(* IEC 61131-3 sources: codesys-framework/txt/application/WeVe IO (library)/Analog Input/FB_AnalogInput, 2 files *)

(* ---- Signals.prop.st ---- *)
PROPERTY Signals : SC_AnalogInputSignals

// --- BEGIN IMPLEMENTATION ---

// ----------- GET -----------
VAR
END_VAR

// -- BEGIN IMPLEMENTATION GET --
Signals := _scSignalValue;

(* ---- SysPar.prop.st ---- *)
PROPERTY SysPar : SC_SystemParametersAnalogInput

// --- BEGIN IMPLEMENTATION ---

// ----------- SET -----------
VAR
END_VAR

// -- BEGIN IMPLEMENTATION SET --
_scSysPar := SysPar;
